	IF InitMqttDone THEN
		pMqttPublishQueue^.AddMessage(
			Payload := REAL_TO_STRING(TOTAL_ACTIVE_ENERGY),
			Topic := CONCAT(CONCAT(MqttPublishTopicPrefix^, MqttPublishTopicSuffix), '/TOTAE' ),
			Qos := MQTT.QoS.ExactlyOnce,
			MqttRetain := FALSE
		);
		pMqttPublishQueue^.AddMessage(
			Payload := REAL_TO_STRING(TOTAL_REACTIVE_ENERGY),
			Topic := CONCAT(CONCAT(MqttPublishTopicPrefix^, MqttPublishTopicSuffix), '/TOTRE' ),
			Qos := MQTT.QoS.ExactlyOnce,
			MqttRetain := FALSE
		);
	END_IF
END_IF
          

METHOD ProcessDataArray
  VAR_INPUT
    Error : POINTER TO BOOL;
    Data : POINTER TO ARRAY[0..124] OF WORD;
  END_VAR
                  IF Error^ THEN
	PubMqttMessage(Suffix := '/availability', Data := 'offline');
ELSE
	PubMqttMessage(Suffix := '/availability', Data := 'online');
END_IF

IF ActiveRtuQuery = 1 THEN
	THIS^.Error1 := Error^;
	THIS^.timerData1.IN := TRUE;
	IF NOT Error^ THEN
		THIS^.VOLTAGE := SwapWordsToReal(Data^[0], Data^[1]);
		THIS^.CURRENT := SwapWordsToReal(Data^[6], Data^[7]);
		THIS^.ACTIVEPOWER := SwapWordsToReal(Data^[12], Data^[13]);
		THIS^.APPARENT_POWER := SwapWordsToReal(Data^[18], Data^[19]);
		THIS^.REACTIVE_POWER := SwapWordsToReal(Data^[24], Data^[25]);
		THIS^.POWER_FACTOR := SwapWordsToReal(Data^[30], Data^[31]);
		THIS^.PHASE_ANGLE := SwapWordsToReal(Data^[36], Data^[37]);
		THIS^.Update1 := TRUE;
	END_IF
ELSIF ActiveRtuQuery = 2 THEN
	THIS^.Error2:= Error^;
	THIS^.timerData2.IN := TRUE;
	IF NOT Error^ THEN		
		THIS^.FREQUENCY := SwapWordsToReal(Data^[0], Data^[1]);
		THIS^.IMPORT_ACTIVE_ENERGY := SwapWordsToReal(Data^[2], Data^[3]);
		THIS^.EXPORT_ACTIVE_ENERGY := SwapWordsToReal(Data^[4], Data^[5]);
		THIS^.IMPORT_REACTIVE_ENERGY := SwapWordsToReal(Data^[6], Data^[7]);
		THIS^.EXPORT_REACTIVE_ENERGY := SwapWordsToReal(Data^[8], Data^[9]);
		THIS^.Update2 := TRUE;
	END_IF
ELSIF ActiveRtuQuery = 3 THEN
	THIS^.Error3 := Error^;
	THIS^.timerData3.IN := TRUE;
	IF NOT Error^ THEN
		THIS^.TOTAL_ACTIVE_ENERGY := SwapWordsToReal(Data^[0], Data^[1]);
		THIS^.TOTAL_REACTIVE_ENERGY := SwapWordsToReal(Data^[2], Data^[3]);
		THIS^.Update3 := TRUE;
	END_IF	
END_IF

ActiveRtuQuery := 0;
ActiveDevice := FALSE;




                
END_METHOD

METHOD InitRS485
  VAR_INPUT
    Data1PollingInterval : TIME;
    Data2PollingInterval : TIME;
    Data3PollingInterval : TIME;
    DeviceAddress : BYTE;
  END_VAR
                  THIS^.timerData1.PT := Data1PollingInterval;
THIS^.timerData2.PT := Data2PollingInterval;
THIS^.timerData3.PT := Data3PollingInterval;

THIS^.Data1RtuQuery.DeviceId := DeviceAddress;
THIS^.Data2RtuQuery.DeviceId := DeviceAddress;
THIS^.Data3RtuQuery.DeviceId := DeviceAddress;

THIS^.timerData1.IN := TRUE;
THIS^.timerData2.IN := TRUE;
THIS^.timerData3.IN := TRUE;

THIS^.InitRS485Done := TRUE;
                
END_METHOD

METHOD InitMqtt
  VAR_INPUT
    MQTTPublishPrefix : POINTER TO STRING;
    pMqttPublishQueue : POINTER TO FB_MqttPublishQueue;
  END_VAR
  VAR
    InstanceNamePt : POINTER TO STRING;
  END_VAR
                  THIS^.pMqttPublishQueue := pMqttPublishQueue;
THIS^.MqttPublishTopicPrefix := MQTTPublishPrefix;

InstanceNamePt := CommonTypesAndFunctions.FindLastDot(ADR(THIS^.InstanceName)) + 1;
THIS^.MqttPublishTopicSuffix := InstanceNamePt^;

THIS^.InitMqttDone := TRUE;
                
END_METHOD

METHOD RequestBusTime : BOOL
                  IF NOT InitRS485Done THEN	
	RequestBusTime := FALSE;	
ELSIF timerData1.Q OR timerData2.Q OR timerData3.Q THEN
	RequestBusTime := TRUE;	
ELSE
	RequestBusTime := FALSE;		
END_IF
                
END_METHOD

METHOD GetRtuQuery : RS485_RtuQuery
                  IF timerData1.Q THEN
	THIS^.timerData1.IN := FALSE;
	THIS^.ActiveRtuQuery := 1;
	GetRtuQuery := THIS^.Data1RtuQuery;
ELSIF timerData2.Q THEN
	THIS^.timerData2.IN := FALSE;
	THIS^.ActiveRtuQuery := 2;
	GetRtuQuery := THIS^.Data2RtuQuery;
ELSIF timerData3.Q THEN
	THIS^.timerData3.IN := FALSE;
	THIS^.ActiveRtuQuery := 3;
	GetRtuQuery := THIS^.Data3RtuQuery;	
END_IF
                
END_METHOD

METHOD PubMqttMessage
  VAR_INPUT
    Suffix : STRING(100);
    Data : STRING(100);
  END_VAR
                  IF InitMqttDone THEN
		pMqttPublishQueue^.AddMessage(
			Payload := Data,
			Topic := CONCAT(CONCAT(MqttPublishTopicPrefix^, MqttPublishTopicSuffix), Suffix ),
			Qos := MQTT.QoS.ExactlyOnce,
			MqttRetain := FALSE
		);
END_IF
                
END_METHOD
END_FUNCTION_BLOCK

{attribute 'reflection'}
FUNCTION_BLOCK FB_RS485_ESERA_1WIRE_GATEWAY_MQTT IMPLEMENTS RS485Device
  VAR
    {attribute 'instance-path'}
    {attribute 'noinit'}
    InstanceName : STRING;  (* object's full instance name *)
    InitRS485Done : BOOL := FALSE;
    DeviceAddress : BYTE;
    OwdDevices : ARRAY[1..30] OF FB_RS485_ESERA_OWD_MQTT;
    ActiveDevice : BOOL := FALSE;
    ActiveOwd : UINT := 0;
    loopCounter : UINT;
    timerData : TON;
  END_VAR

            timerData();

FOR loopCounter := 1 TO 30 DO
	OwdDevices[loopCounter]();
END_FOR
          

METHOD GetRtuQuery : RS485_RtuQuery
                  IF timerData.Q THEN
	THIS^.timerData.IN := FALSE;
	GetRtuQuery := THIS^.OwdDevices[ActiveOwd].GetRtuQuery();	
END_IF
                
END_METHOD

METHOD ProcessDataArray
  VAR_INPUT
    Error : POINTER TO BOOL;
    Data : POINTER TO ARRAY[0..124] OF WORD;
  END_VAR
                  THIS^.OwdDevices[ActiveOwd].ProcessDataArray(
	Data := Data,
	Error := Error
);
THIS^.ActiveOwd := 0;
THIS^.timerData.IN := TRUE;
                
END_METHOD

METHOD RequestBusTime : BOOL
                  IF NOT InitRS485Done OR NOT timerData.Q THEN	
	RequestBusTime := FALSE;
ELSE
	FOR loopCounter := 1 TO 30 DO
		IF OwdDevices[loopCounter].RequestBusTime() AND RequestBusTime = FALSE THEN
			THIS^.ActiveOwd := loopCounter;
			RequestBusTime := TRUE;			
		END_IF
	END_FOR
END_IF
                
END_METHOD

METHOD InitRS485
  VAR_INPUT
    DeviceAddress : BYTE;
  END_VAR
                  THIS^.DeviceAddress := DeviceAddress;
THIS^.timerData.PT := T#250MS;
THIS^.timerData.IN := TRUE;
THIS^.InitRS485Done := TRUE;
                
END_METHOD

METHOD InitMqtt
  VAR_INPUT
    MQTTPublishPrefix : POINTER TO STRING;
    pMqttPublishQueue : POINTER TO FB_MqttPublishQueue;
  END_VAR
  VAR
    InstanceNamePt : POINTER TO STRING;
  END_VAR
                  InstanceNamePt := CommonTypesAndFunctions.FindLastDot(ADR(THIS^.InstanceName)) + 1;

FOR loopCounter := 1 TO 30 DO
		OwdDevices[loopCounter].InitMqtt(
			MQTTPublishPrefix := MQTTPublishPrefix,
			MqttPublishTopicSuffix := InstanceNamePt^,
			pMqttPublishQueue := pMqttPublishQueue
		);
END_FOR
                
END_METHOD

METHOD EnableOwd : BOOL
  VAR_INPUT
    OwdNumber : UINT;
    DataPollingInterval : TIME;
  END_VAR
                  THIS^.OwdDevices[OwdNumber].InitOwd(
	DeviceAddress := THIS^.DeviceAddress,
	OwdNumber := OwdNumber,
	DataPollingInterval := DataPollingInterval
);
                
END_METHOD
END_FUNCTION_BLOCK

FUNCTION_BLOCK FB_RS485_ESERA_OWD_MQTT
  VAR_OUTPUT
    OWD_VOLTAGE : REAL := 0;
    TEMPERATURE : REAL := 0;
    HUMIDITY : REAL := 0;
    DEW_POINT : REAL := 0;
    AIR_QUALITY : REAL := 0;
    BRIGHTNESS : REAL := 0;
    DataAvailable : BOOL := FALSE;
    Error : BOOL := FALSE;
  END_VAR
  VAR
    OwdNumber : UINT;
    InitMqttDone : BOOL;
    MqttPublishTopicPrefix : POINTER TO STRING;
    MqttPublishTopicSuffix : STRING(50);
    pMqttPublishQueue : POINTER TO FB_MqttPublishQueue;
    InitOwdDone : BOOL := FALSE;
    timerData : TON;
    RtuQuery : RS485_RtuQuery := (FunctionCode := 3, ReadAddress := 100, ReadQuantity := 17);
  END_VAR

            timerData();


          

METHOD InitOwd
  VAR_INPUT
    DeviceAddress : BYTE;
    OwdNumber : UINT;
    DataPollingInterval : TIME;
  END_VAR
                  THIS^.RtuQuery.DeviceId := DeviceAddress;
THIS^.RtuQuery.ReadAddress := OwdNumber * 100;
THIS^.timerData.PT := DataPollingInterval;
THIS^.OwdNumber := OwdNumber;

THIS^.timerData.IN := TRUE;

THIS^.InitOwdDone := TRUE;
                
END_METHOD

METHOD InitMqtt
  VAR_INPUT
    MQTTPublishPrefix : POINTER TO STRING;
    MqttPublishTopicSuffix : STRING(255);
    pMqttPublishQueue : POINTER TO FB_MqttPublishQueue;
  END_VAR
                  THIS^.MqttPublishTopicPrefix := MQTTPublishPrefix;
THIS^.MqttPublishTopicSuffix := MqttPublishTopicSuffix;
THIS^.pMqttPublishQueue := pMqttPublishQueue;

THIS^.InitMqttDone := TRUE;
                
END_METHOD

METHOD PubMqttMessage
  VAR_INPUT
    Suffix : STRING(100);
    Data : STRING(100);
  END_VAR
                  IF InitMqttDone THEN
		pMqttPublishQueue^.AddMessage(
			Payload := Data,
			Topic := CONCAT(CONCAT(CONCAT(CONCAT(MqttPublishTopicPrefix^, MqttPublishTopicSuffix), '/OWD/'), UINT_TO_STRING(OwdNumber)), Suffix ),
			Qos := MQTT.QoS.ExactlyOnce,
			MqttRetain := FALSE
		);
END_IF
                
END_METHOD

METHOD ProcessTemperature
  VAR_INPUT
    Data : WORD;
  END_VAR
                  THIS^.TEMPERATURE := WORD_TO_REAL(Data) / 100;
PubMqttMessage(Suffix := '/TEMP', Data := REAL_TO_STRING(TEMPERATURE));
                
END_METHOD

METHOD ProcessOwdVoltage
  VAR_INPUT
    Data : WORD;
  END_VAR
                  THIS^.OWD_VOLTAGE := WORD_TO_REAL(Data) / 100;
PubMqttMessage(Suffix := '/OWDV', Data := REAL_TO_STRING(OWD_VOLTAGE));
                
END_METHOD

METHOD ProcessHumidity
  VAR_INPUT
    Data : WORD;
  END_VAR
                  THIS^.HUMIDITY := WORD_TO_REAL(Data) / 100;
PubMqttMessage(Suffix := '/HUM', Data := REAL_TO_STRING(HUMIDITY));
                
END_METHOD

METHOD ProcessDewPoint
  VAR_INPUT
    Data : WORD;
  END_VAR
                  THIS^.DEW_POINT := WORD_TO_REAL(Data) / 100;
PubMqttMessage(Suffix := '/DEWP', Data := REAL_TO_STRING(DEW_POINT));
                
END_METHOD

METHOD ProcessAirQuality
  VAR_INPUT
    Data : WORD;
  END_VAR
                  THIS^.AIR_QUALITY := WORD_TO_REAL(Data) / 100;
PubMqttMessage(Suffix := '/AIRQ', Data := REAL_TO_STRING(AIR_QUALITY));
                
END_METHOD

METHOD GetRtuQuery : RS485_RtuQuery
                  IF timerData.Q THEN
	THIS^.timerData.IN := FALSE;
	GetRtuQuery := THIS^.RtuQuery;	
END_IF
                
END_METHOD

METHOD ProcessDataArray
  VAR_INPUT
    Error : POINTER TO BOOL;
    Data : POINTER TO ARRAY[0..124] OF WORD;
  END_VAR
                  THIS^.timerData.IN := TRUE;

IF WORD_TO_INT(Data^[12]) <> 0 OR Error^ THEN
	THIS^.Error := TRUE;
	PubMqttMessage(Suffix := '/availability', Data := 'offline');
ELSE 	
	THIS^.Error := FALSE;
	THIS^.DataAvailable := TRUE;
	PubMqttMessage(Suffix := '/availability', Data := 'online');
END_IF

// Data handling
IF NOT Error^ AND WORD_TO_INT(Data^[12]) = 0 THEN
	IF Data^[16] = 11151 OR Data^[16] = 11152 THEN // Temperature, humidity & air quality
		ProcessTemperature(Data^[0]);		
		ProcessOwdVoltage(Data^[2]);
		ProcessHumidity(Data^[4]);
		ProcessDewPoint(Data^[6]);
		ProcessAirQuality(Data^[8]);
	ELSIF Data^[16] = 11102 OR Data^[16] = 11113 OR Data^[16] = 11120 OR Data^[16] = 11148 OR Data^[16] = 11150 OR Data^[16] = 11160 THEN // Temperature, humidity
		ProcessTemperature(Data^[0]);		
		ProcessOwdVoltage(Data^[2]);
		ProcessHumidity(Data^[4]);
		ProcessDewPoint(Data^[6]);
	ELSIF Data^[16] = 11121 OR Data^[16] = 11132 OR Data^[16] = 11134 OR Data^[16] = 11135 THEN // Temperature, humidity, brightness
		ProcessTemperature(Data^[0]);		
		ProcessOwdVoltage(Data^[2]);
		ProcessHumidity(Data^[4]);
		ProcessDewPoint(Data^[6]);
		ProcessBrigthness(Data^[8]);
	ELSIF Data^[16] = 1820  THEN // Temperature DS18B20
        ProcessTemperature(Data^[0]);
	END_IF		
END_IF
                
END_METHOD

METHOD RequestBusTime : BOOL
                  IF NOT InitOwdDone THEN	
	RequestBusTime := FALSE;	
ELSIF timerData.Q THEN
	RequestBusTime := TRUE;
ELSE
	RequestBusTime := FALSE;	
END_IF
                
END_METHOD

METHOD ProcessBrigthness
  VAR_INPUT
    Data : WORD;
  END_VAR
                  THIS^.BRIGHTNESS := WORD_TO_REAL(Data) / 100;
PubMqttMessage(Suffix := '/BNESS', Data := REAL_TO_STRING(BRIGHTNESS));
                
END_METHOD
END_FUNCTION_BLOCK

{attribute 'reflection'}
FUNCTION_BLOCK FB_VIRTUAL_BOOL_MQTT EXTENDS FB_MQTT_BASE IMPLEMENTS MQTT.MQTT_SUBSCRIBE_CALLBACK
  VAR_INPUT
    IN : BOOL;
  END_VAR
  VAR_OUTPUT
    OUT : BOOL;
  END_VAR
  VAR
    {attribute 'instance-path'}
    {attribute 'noinit'}
    InstancePath : STRING;  (* Refelection: object's full instance name *)
    Startup : BOOL := TRUE;
    UpdateFlag : BOOL;
    VirtualMode : VIRTUAL_MODES;
    DefaultValue : BOOL;
    SetDefaultValueStartup : BOOL;
    PublishAtStartup : BOOL;
    UsePersistentAtStartup : BOOL;
    ConfirmReceival : BOOL;
    MqttMessageReceived : BOOL;
    PreviousIn : BOOL;
  END_VAR
  VAR PERSISTENT
    PreviousState : BOOL;  (* To retain output state through powercycles *)
  END_VAR

            IF VirtualMode = VIRTUAL_MODES.Output THEN
	IF (Startup AND PublishAtStartup) OR (UpdateFlag OR IN <> PreviousIn) AND InitMqttDone THEN
	pMqttPublishQueue^.AddMessage(
		Payload := BOOL_TO_STRING(IN),
		Topic := CONCAT(MqttPublishTopicPrefix^, MqttPublishTopicSuffix),
		Qos := MqttQos,
		MqttRetain := MqttRetain
	);
	Startup:=FALSE;
	UpdateFlag := FALSE;
	PreviousIn := IN;
	END_IF
ELSIF VirtualMode = VIRTUAL_MODES.Input THEN
	IF Startup AND SetDefaultValueStartup THEN
		OUT := DefaultValue;
	ELSIF UsePersistentAtStartup THEN
		OUT := PreviousState;
	END_IF	
	
	IF ((Startup AND PublishAtStartup) OR (ConfirmReceival AND MqttMessageReceived)) AND InitMqttDone THEN
	pMqttPublishQueue^.AddMessage(
		Payload := BOOL_TO_STRING(OUT),
		Topic := CONCAT(MqttPublishTopicPrefix^, MqttPublishTopicSuffix),
		Qos := MqttQos,
		MqttRetain := MqttRetain
	);
	Startup:=FALSE;
	MqttMessageReceived := FALSE;
	PreviousState:=OUT;
	END_IF		
	
END_IF
          

METHOD InitMqtt
  VAR_INPUT
    MQTTPublishPrefix : POINTER TO STRING;
    MQTTSubscribePrefix : POINTER TO STRING;
    pMqttPublishQueue : POINTER TO FB_MqttPublishQueue;
    pMqttCallbackCollector : POINTER TO MQTT.CallbackCollector;
    MqttQos : MQTT.QoS;
    MqttRetain : BOOL;
  END_VAR
                  InitMqttDone := TRUE;

SUPER^._InstancePath := THIS^.InstancePath; // Due to reflection its location is important

(*pass trough*)
THIS^.pMqttPublishQueue := pMqttPublishQueue;
THIS^.MqttPublishTopicPrefix:=MQTTPublishPrefix;
THIS^.MQTTSubscribeTopicPrefix:=MQTTSubscribePrefix;
THIS^.pMqttPublishQueue:=pMqttPublishQueue;
THIS^.MqttQos:=MqttQos;
THIS^.MqttRetain:=MqttRetain;


SUPER^.InitBaseMqtt();
pMqttCallbackCollector^.put(instance:= THIS^); // register the FB agains the collector so mqtt events can be received


                
END_METHOD

METHOD PublishReceived : BOOL
  VAR_INPUT
    Data : MQTT.CALLBACK_DATA;  (* Collection of recived Data *)
  END_VAR
                  //first check if Mqtt is initialized and FB in input mode, otherwise do nothing
IF NOT(InitMqttDone) AND VirtualMode <> VIRTUAL_MODES.Input THEN
	//mark the interface call from the collector as done
	PublishReceived := TRUE;
//check if the packet is for this FB
ELSIF CommonTypesAndFunctions.StrEquals(str1:= ADR(MQTTSubscribeTopic), str2:= Data.TopicOut) THEN
	//mark the interface call from the collector as done
	PublishReceived := TRUE;
	//process the data
	IF CommonTypesAndFunctions.StrEquals(str1:= Data.PayloadString, str2:= ADR('TRUE')) THEN
		THIS^.OUT := TRUE;
		MqttMessageReceived := TRUE;
	END_IF
	IF CommonTypesAndFunctions.StrEquals(str1:= Data.PayloadString, str2:= ADR('FALSE')) THEN
		THIS^.OUT := FALSE;
		MqttMessageReceived := TRUE;
	END_IF
END_IF 
                
END_METHOD

METHOD ConfigureFunctionBlockAsVirtualInput : BOOL
  VAR_INPUT
    DefaultValue : BOOL;
    SetDefaultValueStartup : BOOL;
    PublishAtStartup : BOOL;
    UsePersistentAtStartup : BOOL;
    ConfirmReceival : BOOL;
  END_VAR
                  THIS^.DefaultValue:=DefaultValue;
THIS^.SetDefaultValueStartup:=SetDefaultValueStartup;
THIS^.PublishAtStartup:=PublishAtStartup;
THIS^.UsePersistentAtStartup:=UsePersistentAtStartup;
THIS^.ConfirmReceival:=ConfirmReceival;
THIS^.VirtualMode:=VIRTUAL_MODES.Input;
                
END_METHOD

METHOD SetValue : BOOL
  VAR_INPUT
    Value : BOOL;
  END_VAR
                  THIS^.OUT:=Value;
THIS^.UpdateFlag:=TRUE;
                
END_METHOD

METHOD ConfigureFunctionBlockAsVirtualOutput : BOOL
  VAR_INPUT
    PublishAtStartup : BOOL;
  END_VAR
                  THIS^.PublishAtStartup:=PublishAtStartup;
THIS^.VirtualMode:=VIRTUAL_MODES.Output;
                
END_METHOD
END_FUNCTION_BLOCK

{attribute 'reflection'}
FUNCTION_BLOCK FB_VIRTUAL_INT_MQTT EXTENDS FB_MQTT_BASE IMPLEMENTS MQTT.MQTT_SUBSCRIBE_CALLBACK
  VAR_INPUT
    IN : INT;
  END_VAR
  VAR_OUTPUT
    OUT : INT;
  END_VAR
  VAR
    {attribute 'instance-path'}
    {attribute 'noinit'}
    InstancePath : STRING;  (* Refelection: object's full instance name *)
    Startup : BOOL := TRUE;
    UpdateFlag : BOOL;
    VirtualMode : VIRTUAL_MODES;
    DefaultValue : INT;
    SetDefaultValueStartup : BOOL;
    PublishAtStartup : BOOL;
    UsePersistentAtStartup : BOOL;
    ConfirmReceival : BOOL;
    MqttMessageReceived : BOOL;
    PreviousIn : INT;
  END_VAR
  VAR PERSISTENT
    PreviousState : INT;  (* To retain output state through powercycles *)
  END_VAR

            IF VirtualMode = VIRTUAL_MODES.Output THEN
	IF (Startup AND PublishAtStartup) OR (UpdateFlag OR IN <> PreviousIn) AND InitMqttDone THEN
	pMqttPublishQueue^.AddMessage(
		Payload := INT_TO_STRING(IN),
		Topic := CONCAT(MqttPublishTopicPrefix^, MqttPublishTopicSuffix),
		Qos := MqttQos,
		MqttRetain := MqttRetain
	);
	Startup:=FALSE;
	UpdateFlag := FALSE;
	PreviousIn := IN;
	END_IF
ELSIF VirtualMode = VIRTUAL_MODES.Input THEN
	IF Startup AND SetDefaultValueStartup THEN
		OUT := DefaultValue;
	ELSIF UsePersistentAtStartup THEN
		OUT := PreviousState;
	END_IF	
	
	IF ((Startup AND PublishAtStartup) OR (ConfirmReceival AND MqttMessageReceived)) AND InitMqttDone THEN
	pMqttPublishQueue^.AddMessage(
		Payload := INT_TO_STRING(OUT),
		Topic := CONCAT(MqttPublishTopicPrefix^, MqttPublishTopicSuffix),
		Qos := MqttQos,
		MqttRetain := MqttRetain
	);
	Startup:=FALSE;
	MqttMessageReceived := FALSE;
	PreviousState:=OUT;
	END_IF		
	
END_IF
          

METHOD ConfigureFunctionBlockAsVirtualOutput : BOOL
  VAR_INPUT
    PublishAtStartup : BOOL;
  END_VAR
                  THIS^.PublishAtStartup:=PublishAtStartup;
THIS^.VirtualMode:=VIRTUAL_MODES.Output;
                
END_METHOD

METHOD InitMqtt
  VAR_INPUT
    MQTTPublishPrefix : POINTER TO STRING;
    MQTTSubscribePrefix : POINTER TO STRING;
    pMqttPublishQueue : POINTER TO FB_MqttPublishQueue;
    pMqttCallbackCollector : POINTER TO MQTT.CallbackCollector;
    MqttQos : MQTT.QoS;
    MqttRetain : BOOL;
  END_VAR
                  InitMqttDone := TRUE;

SUPER^._InstancePath := THIS^.InstancePath; // Due to reflection its location is important

(*pass trough*)
THIS^.pMqttPublishQueue := pMqttPublishQueue;
THIS^.MqttPublishTopicPrefix:=MQTTPublishPrefix;
THIS^.MQTTSubscribeTopicPrefix:=MQTTSubscribePrefix;
THIS^.pMqttPublishQueue:=pMqttPublishQueue;
THIS^.MqttQos:=MqttQos;
THIS^.MqttRetain:=MqttRetain;


SUPER^.InitBaseMqtt();
pMqttCallbackCollector^.put(instance:= THIS^); // register the FB agains the collector so mqtt events can be received


                
END_METHOD

METHOD PublishReceived : BOOL
  VAR_INPUT
    Data : MQTT.CALLBACK_DATA;  (* Collection of recived Data *)
  END_VAR
                  //first check if Mqtt is initialized and FB in input mode, otherwise do nothing
IF NOT(InitMqttDone) AND VirtualMode <> VIRTUAL_MODES.Input THEN
	//mark the interface call from the collector as done
	PublishReceived := TRUE;
//check if the packet is for this FB
ELSIF CommonTypesAndFunctions.StrEquals(str1:= ADR(MQTTSubscribeTopic), str2:= Data.TopicOut) THEN
	//mark the interface call from the collector as done
	PublishReceived := TRUE;
	//process the data
	IF OSCAT_BASIC.IS_NUM(str:= Data.PayloadString^) THEN
		THIS^.OUT := STRING_TO_INT(Data.PayloadString^);	
		MqttMessageReceived := TRUE;	
	END_IF
END_IF 
                
END_METHOD

METHOD ConfigureFunctionBlockAsVirtualInput : BOOL
  VAR_INPUT
    DefaultValue : INT;
    SetDefaultValueStartup : BOOL;
    PublishAtStartup : BOOL;
    UsePersistentAtStartup : BOOL;
    ConfirmReceival : BOOL;
  END_VAR
                  THIS^.DefaultValue:=DefaultValue;
THIS^.SetDefaultValueStartup:=SetDefaultValueStartup;
THIS^.PublishAtStartup:=PublishAtStartup;
THIS^.UsePersistentAtStartup:=UsePersistentAtStartup;
THIS^.ConfirmReceival:=ConfirmReceival;
THIS^.VirtualMode:=VIRTUAL_MODES.Input;
                
END_METHOD

METHOD SetValue : BOOL
  VAR_INPUT
    Value : INT;
  END_VAR
                  THIS^.OUT:=Value;
THIS^.UpdateFlag:=TRUE;
                
END_METHOD
END_FUNCTION_BLOCK

{attribute 'reflection'}
FUNCTION_BLOCK FB_VIRTUAL_REAL_MQTT EXTENDS FB_MQTT_BASE IMPLEMENTS MQTT.MQTT_SUBSCRIBE_CALLBACK
  VAR_INPUT
    IN : REAL;
  END_VAR
  VAR_OUTPUT
    OUT : REAL;
  END_VAR
  VAR
    {attribute 'instance-path'}
    {attribute 'noinit'}
    InstancePath : STRING;  (* Refelection: object's full instance name *)
    Startup : BOOL := TRUE;
    UpdateFlag : BOOL;
    VirtualMode : VIRTUAL_MODES;
    DefaultValue : REAL;
    SetDefaultValueStartup : BOOL;
    PublishAtStartup : BOOL;
    UsePersistentAtStartup : BOOL;
    ConfirmReceival : BOOL;
    MqttMessageReceived : BOOL;
    PreviousIn : REAL;
  END_VAR
  VAR PERSISTENT
    PreviousState : REAL;  (* To retain output state through powercycles *)
  END_VAR

            IF VirtualMode = VIRTUAL_MODES.Output THEN
	IF (Startup AND PublishAtStartup) OR (UpdateFlag OR IN <> PreviousIn) AND InitMqttDone THEN
	pMqttPublishQueue^.AddMessage(
		Payload := REAL_TO_STRING(IN),
		Topic := CONCAT(MqttPublishTopicPrefix^, MqttPublishTopicSuffix),
		Qos := MqttQos,
		MqttRetain := MqttRetain
	);
	Startup:=FALSE;
	UpdateFlag := FALSE;
	PreviousIn := IN;
	END_IF
ELSIF VirtualMode = VIRTUAL_MODES.Input THEN
	IF Startup AND SetDefaultValueStartup THEN
		OUT := DefaultValue;
	ELSIF UsePersistentAtStartup THEN
		OUT := PreviousState;
	END_IF	
	
	IF ((Startup AND PublishAtStartup) OR (ConfirmReceival AND MqttMessageReceived)) AND InitMqttDone THEN
	pMqttPublishQueue^.AddMessage(
		Payload := REAL_TO_STRING(OUT),
		Topic := CONCAT(MqttPublishTopicPrefix^, MqttPublishTopicSuffix),
		Qos := MqttQos,
		MqttRetain := MqttRetain
	);
	Startup:=FALSE;
	MqttMessageReceived := FALSE;
	PreviousState:=OUT;
	END_IF		
	
END_IF
          

METHOD ConfigureFunctionBlockAsVirtualOutput : BOOL
  VAR_INPUT
    PublishAtStartup : BOOL;
  END_VAR
                  THIS^.PublishAtStartup:=PublishAtStartup;
THIS^.VirtualMode:=VIRTUAL_MODES.Output;
                
END_METHOD

METHOD InitMqtt
  VAR_INPUT
    MQTTPublishPrefix : POINTER TO STRING;
    MQTTSubscribePrefix : POINTER TO STRING;
    pMqttPublishQueue : POINTER TO FB_MqttPublishQueue;
    pMqttCallbackCollector : POINTER TO MQTT.CallbackCollector;
    MqttQos : MQTT.QoS;
    MqttRetain : BOOL;
  END_VAR
                  InitMqttDone := TRUE;

SUPER^._InstancePath := THIS^.InstancePath; // Due to reflection its location is important

(*pass trough*)
THIS^.pMqttPublishQueue := pMqttPublishQueue;
THIS^.MqttPublishTopicPrefix:=MQTTPublishPrefix;
THIS^.MQTTSubscribeTopicPrefix:=MQTTSubscribePrefix;
THIS^.pMqttPublishQueue:=pMqttPublishQueue;
THIS^.MqttQos:=MqttQos;
THIS^.MqttRetain:=MqttRetain;


SUPER^.InitBaseMqtt();
pMqttCallbackCollector^.put(instance:= THIS^); // register the FB agains the collector so mqtt events can be received


                
END_METHOD

METHOD PublishReceived : BOOL
  VAR_INPUT
    Data : MQTT.CALLBACK_DATA;  (* Collection of recived Data *)
  END_VAR
                  //first check if Mqtt is initialized and FB in input mode, otherwise do nothing
IF NOT(InitMqttDone) AND VirtualMode <> VIRTUAL_MODES.Input THEN
	//mark the interface call from the collector as done
	PublishReceived := TRUE;
//check if the packet is for this FB
ELSIF CommonTypesAndFunctions.StrEquals(str1:= ADR(MQTTSubscribeTopic), str2:= Data.TopicOut) THEN
	//mark the interface call from the collector as done
	PublishReceived := TRUE;
	//process the data
	THIS^.OUT := STRING_TO_REAL(Data.PayloadString^);	
	MqttMessageReceived := TRUE;	
END_IF 
                
END_METHOD

METHOD ConfigureFunctionBlockAsVirtualInput : BOOL
  VAR_INPUT
    DefaultValue : REAL;
    SetDefaultValueStartup : BOOL;
    PublishAtStartup : BOOL;
    UsePersistentAtStartup : BOOL;
    ConfirmReceival : BOOL;
  END_VAR
                  THIS^.DefaultValue:=DefaultValue;
THIS^.SetDefaultValueStartup:=SetDefaultValueStartup;
THIS^.PublishAtStartup:=PublishAtStartup;
THIS^.UsePersistentAtStartup:=UsePersistentAtStartup;
THIS^.ConfirmReceival:=ConfirmReceival;
THIS^.VirtualMode:=VIRTUAL_MODES.Input;
                
END_METHOD

METHOD SetValue : BOOL
  VAR_INPUT
    Value : REAL;
  END_VAR
                  THIS^.OUT:=Value;
THIS^.UpdateFlag:=TRUE;
                
END_METHOD
END_FUNCTION_BLOCK

{attribute 'reflection'}
FUNCTION_BLOCK FB_VIRTUAL_STRING_MQTT EXTENDS FB_MQTT_BASE IMPLEMENTS MQTT.MQTT_SUBSCRIBE_CALLBACK
  VAR_INPUT
    IN : STRING;
  END_VAR
  VAR_OUTPUT
    OUT : STRING;
  END_VAR
  VAR
    {attribute 'instance-path'}
    {attribute 'noinit'}
    InstancePath : STRING;  (* Refelection: object's full instance name *)
    Startup : BOOL := TRUE;
    UpdateFlag : BOOL;
    VirtualMode : VIRTUAL_MODES;
    DefaultValue : STRING;
    SetDefaultValueStartup : BOOL;
    PublishAtStartup : BOOL;
    UsePersistentAtStartup : BOOL;
    ConfirmReceival : BOOL;
    MqttMessageReceived : BOOL;
    PreviousIn : STRING;
  END_VAR
  VAR PERSISTENT
    PreviousState : STRING;  (* To retain output state through powercycles *)
  END_VAR

            IF VirtualMode = VIRTUAL_MODES.Output THEN
	IF (Startup AND PublishAtStartup) OR (UpdateFlag OR IN <> PreviousIn) AND InitMqttDone THEN
	pMqttPublishQueue^.AddMessage(
		Payload := IN,
		Topic := CONCAT(MqttPublishTopicPrefix^, MqttPublishTopicSuffix),
		Qos := MqttQos,
		MqttRetain := MqttRetain
	);
	Startup:=FALSE;
	UpdateFlag := FALSE;
	PreviousIn := IN;
	END_IF
ELSIF VirtualMode = VIRTUAL_MODES.Input THEN
	IF Startup AND SetDefaultValueStartup THEN
		OUT := DefaultValue;
	ELSIF UsePersistentAtStartup THEN
		OUT := PreviousState;
	END_IF	
	
	IF ((Startup AND PublishAtStartup) OR (ConfirmReceival AND MqttMessageReceived)) AND InitMqttDone THEN
	pMqttPublishQueue^.AddMessage(
		Payload := OUT,
		Topic := CONCAT(MqttPublishTopicPrefix^, MqttPublishTopicSuffix),
		Qos := MqttQos,
		MqttRetain := MqttRetain
	);
	Startup:=FALSE;
	MqttMessageReceived := FALSE;
	PreviousState:=OUT;
	END_IF		
	
END_IF
          

METHOD InitMqtt
  VAR_INPUT
    MQTTPublishPrefix : POINTER TO STRING;
    MQTTSubscribePrefix : POINTER TO STRING;
    pMqttPublishQueue : POINTER TO FB_MqttPublishQueue;
    pMqttCallbackCollector : POINTER TO MQTT.CallbackCollector;
    MqttQos : MQTT.QoS;
    MqttRetain : BOOL;
  END_VAR
                  InitMqttDone := TRUE;

SUPER^._InstancePath := THIS^.InstancePath; // Due to reflection its location is important

(*pass trough*)
THIS^.pMqttPublishQueue := pMqttPublishQueue;
THIS^.MqttPublishTopicPrefix:=MQTTPublishPrefix;
THIS^.MQTTSubscribeTopicPrefix:=MQTTSubscribePrefix;
THIS^.pMqttPublishQueue:=pMqttPublishQueue;
THIS^.MqttQos:=MqttQos;
THIS^.MqttRetain:=MqttRetain;


SUPER^.InitBaseMqtt();
pMqttCallbackCollector^.put(instance:= THIS^); // register the FB agains the collector so mqtt events can be received


                
END_METHOD

METHOD PublishReceived : BOOL
  VAR_INPUT
    Data : MQTT.CALLBACK_DATA;  (* Collection of recived Data *)
  END_VAR
                  //first check if Mqtt is initialized and FB in input mode, otherwise do nothing
IF NOT(InitMqttDone) AND VirtualMode <> VIRTUAL_MODES.Input THEN
	//mark the interface call from the collector as done
	PublishReceived := TRUE;
//check if the packet is for this FB
ELSIF CommonTypesAndFunctions.StrEquals(str1:= ADR(MQTTSubscribeTopic), str2:= Data.TopicOut) THEN
	//mark the interface call from the collector as done
	PublishReceived := TRUE;
	//process the data
	THIS^.OUT := Data.PayloadString^;	
	MqttMessageReceived := TRUE;
END_IF 
                
END_METHOD

METHOD ConfigureFunctionBlockAsVirtualInput : BOOL
  VAR_INPUT
    DefaultValue : STRING;
    SetDefaultValueStartup : BOOL;
    PublishAtStartup : BOOL;
    UsePersistentAtStartup : BOOL;
    ConfirmReceival : BOOL;
  END_VAR
                  THIS^.DefaultValue:=DefaultValue;
THIS^.SetDefaultValueStartup:=SetDefaultValueStartup;
THIS^.PublishAtStartup:=PublishAtStartup;
THIS^.UsePersistentAtStartup:=UsePersistentAtStartup;
THIS^.ConfirmReceival:=ConfirmReceival;
THIS^.VirtualMode:=VIRTUAL_MODES.Input;
                
END_METHOD

METHOD SetValue : BOOL
  VAR_INPUT
    Value : STRING;
  END_VAR
                  THIS^.OUT:=Value;
THIS^.UpdateFlag:=TRUE;
                
END_METHOD

METHOD ConfigureFunctionBlockAsVirtualOutput : BOOL
  VAR_INPUT
    PublishAtStartup : BOOL;
  END_VAR
                  THIS^.PublishAtStartup:=PublishAtStartup;
THIS^.VirtualMode:=VIRTUAL_MODES.Output;
                
END_METHOD
END_FUNCTION_BLOCK

FUNCTION SwapWordsToReal : REAL
  VAR_INPUT
    wHi : WORD;
    wLo : WORD;
  END_VAR
  VAR
    dwVar : DWORD;
    pt_REAL : POINTER TO REAL;
  END_VAR

            dwVar := SHL(WORD_TO_DWORD(wHi),16) OR WORD_TO_DWORD(wLo);
pt_REAL := ADR(dwVar);
SwapWordsToReal := pt_REAL^;
          
END_FUNCTION

PROGRAM PLC_PRG_MAIN
  VAR
    PLC_Device : FB_PLC_MQTT_DISCOVERY_DEVICE;  (* HOME ASSISTANT DISCOVERY VIA MQTT *)
    FB_DI_PB_001 : FB_INPUT_PUSHBUTTON_MQTT;  (* INPUT FUNCTION BLOCKS *)
    FB_DI_PB_002 : FB_INPUT_PUSHBUTTON_DIMMER_MQTT;
    FB_DO_BIN_001 : FB_OUTPUT_BINARY_MQTT;  (* OUTPUT FUNCTION BLOCKS *)
    FB_DO_BISTABLE_001 : FB_OUTPUT_BISTABLE_MQTT;
    FB_DO_COVER_001 : FB_OUTPUT_COVER_MQTT;  (* COVER FUNCTION BLOCKS *)
    FB_AO_DIMMER_001 : FB_OUTPUT_DIMMER_MQTT;  (* DIMMER FUNCTION BLOCKS *)
    TestOUT : WORD;
    FB_VIRTUAL_INT_001 : FB_VIRTUAL_INT_MQTT;  (* VIRTUAL FUNCTION BLOCKS *)
    FB_VIRTUAL_BOOL_001 : FB_VIRTUAL_BOOL_MQTT;
    FB_VIRTUAL_STRING_001 : FB_VIRTUAL_STRING_MQTT;
    FB_VIRTUAL_REAL_001 : FB_VIRTUAL_REAL_MQTT;
  END_VAR

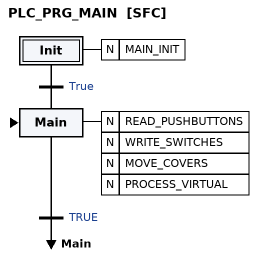
INITIAL_STEP Init:
  MAIN_INIT(N);
END_STEP
TRANSITION FROM Init TO Main
  := True;
END_TRANSITION
STEP Main:
  READ_PUSHBUTTONS(N);
  WRITE_SWITCHES(N);
  MOVE_COVERS(N);
  PROCESS_VIRTUAL(N);
END_STEP
TRANSITION FROM Main TO Main
  := TRUE;
END_TRANSITION

ACTION READ_PUSHBUTTONS:
                      FB_DI_PB_001(PB:= DI_001); (* Provide the input FB the correct phyical input to validate each cyclus *)
FB_DI_PB_002(PB:= DI_002);
                    
END_ACTION

ACTION WRITE_SWITCHES:
                      FB_DO_BIN_001(OUT	=>		DO_001,										(* couple the function block to the physical output *)
	PRIO_HIGH				:=FALSE,  									(* brings the output high regardless of other input values *)
	PRIO_LOW				:=FALSE, 									(* brings the output low regardless of other input values. NOTE: PRIO_HIGH overrules PRIO_LOW input *)
	TOGGLE					:=FB_DI_PB_001.SINGLE 						(* for toggling the output *)	
);

FB_AO_DIMMER_001(
	SINGLE:=FB_DI_PB_001.SINGLE,
	LONG:=FB_DI_PB_001.LONG, 
	P_LONG:=FB_DI_PB_001.P_LONG, 
	Q_OUT => TestOUT,
	SET:=  FB_DI_PB_001.DOUBLE,
	VAL:=125
);

FB_DO_BISTABLE_001();
                    
END_ACTION

ACTION MAIN_INIT:
                      (* MQTT Discovery device*)
PLC_Device.initPlcDevice(
	MqttDiscoveryPrefix := MqttVariables.MqttHADiscoveryPrefix,
	pMqttPublishQueue := ADR(MqttVariables.fbMqttPublishQueue),
	availabilityTopic := MqttVariables.MqttAvailabilityTopic,
	availabilityOnline := MqttVariables.MqttAvailabilityOnlinePayload,
	availabilityOffline := MqttVariables.MqttAvailabilityOfflinePayload
);

(* MQTT logger*)
MqttVariables.MQTT_logger.InitMqtt(
	MQTTPublishPrefix:= ADR(MqttVariables.MqttPubLogPrefix),											
	pMqttPublishQueue := ADR(MqttVariables.fbMqttPublishQueue),				
	MqttQos:=MQTT.QoS.ExactlyOnce, 
	MqttRetain:=FALSE											
);
MqttVariables.MQTT_logger.InitMqttDiscovery(
	Device := ADR(PLC_Device),							(* The device show in Home Assistant *)
);


(* INIT DIGITAL INPUT STUFF *)
FB_DI_PB_001.InitMqtt(
	MQTTPublishPrefix:= ADR(MqttVariables.MqttPushbuttonPrefix),	(* pointer to string prefix for the mqtt publish topic *)
	pMqttPublishQueue := ADR(MqttVariables.fbMqttPublishQueue)		(* pointer to MqttPublishQueue to send a new Mqtt event *)
);

FB_DI_PB_001.InitMqttDiscovery(
	name := 'Button number 001',						(* The name show in Home Assistant frond-end*)
	Device := ADR(PLC_Device),							(* The device show in Home Assistant *)
);

FB_DI_PB_002.InitMqtt(
	MQTTPublishPrefix:= ADR(MqttVariables.MqttPushbuttonPrefix),	
	pMqttPublishQueue := ADR(MqttVariables.fbMqttPublishQueue),
    TRUE,                                                               (* specify whether dimmer value should be outputted on MQTT topic *)
    MQTT.QoS.ExactlyOnce,                                            (* specify the QoS for the dimmer mqtt events (values 0-255) *)    
    5                                                                   (* specify the resolution for the dimmer mqtt events *)    
);


(* ALTER THE DIMMER OUTPUT DEFAULT BEHAVIOR *)
FB_AO_DIMMER_001.ConfigureFunctionBlock(
	T_Debounce:=T#10MS,
	T_Reconfig:=T#10S,
	T_On_Max:=T#0S,
	T_Dimm_Start:=T#400MS,
	T_Dimm:=T#3S,
	Min_On:=50,
	Max_On:=255,
	Soft_Dimm:=TRUE,
	Rst_Out:=FALSE,
	OUT_LinearScaleMin:=11000,
	OUT_LinearScaleMax:=32767
);

(* INIT DMX / ART-NET OUTPUT, OPTIONAL*)
FB_AO_DIMMER_001.InitDmx(
	DmxChannel := 1,							(* The channel *)
	DmxWidth:=1, 								(* Width of DMX channel, 1 or 2, aka 8 or 16 bit *)
	pDmxValues := ADR(DMXVariables.DMX.BUFFER), (* pointer to network buffer *)
	DmxUniverse:=1								(* Universe, but the buffer desides, this is only meta data that ends up in MQTT*)
);

(* INIT HOME ASSISTANT DISCOVERTY*)
FB_AO_DIMMER_001.InitMqttDiscovery(
	name := '001. Office strip cold',					(* The name show in Home Assistant frond-end*)
	Device := ADR(PLC_Device),							(* The device show in Home Assistant *)
);


(* INIT DIGITAL OUTPUT STUFF *)
FB_DO_BISTABLE_001.InitMqtt(
	MQTTPublishPrefix:= ADR(MqttVariables.MqttPubSwitchPrefix),					(* pointer to string prefix for the mqtt publish topic *)
	MQTTSubscribePrefix:= ADR(MqttVariables.MqttSubSwitchPrefix),				(* pointer to string prefix for the mqtt subscribe topic *)
	pMqttPublishQueue := ADR(MqttVariables.fbMqttPublishQueue),					(* pointer to MqttPublishQueue to send a new Mqtt event *)
	pMqttCallbackCollector := ADR(MqttVariables.collector_FB_OUTPUT_SWITCH_MQTT)(* pointer to CallbackCollector to receive Mqtt subscription events *)
);

FB_DO_BISTABLE_001.InitMqttDiscoveryAsLight(
	name := 'light number 1',						(* The name show in Home Assistant frond-end*)
	Device := ADR(PLC_Device),							(* The device show in Home Assistant *)
);

FB_DO_BIN_001.InitMqtt(
	MQTTPublishPrefix:= ADR(MqttVariables.MqttPubSwitchPrefix),					(* pointer to string prefix for the mqtt publish topic *)
	MQTTSubscribePrefix:= ADR(MqttVariables.MqttSubSwitchPrefix),				(* pointer to string prefix for the mqtt subscribe topic *)
	pMqttPublishQueue := ADR(MqttVariables.fbMqttPublishQueue),					(* pointer to MqttPublishQueue to send a new Mqtt event *)
	pMqttCallbackCollector := ADR(MqttVariables.collector_FB_OUTPUT_SWITCH_MQTT)(* pointer to CallbackCollector to receive Mqtt subscription events *)
);

FB_DO_BIN_001.InitMqttDiscoveryAsLight(
	name := 'light number 2',						(* The name show in Home Assistant frond-end*)
	Device := ADR(PLC_Device),							(* The device show in Home Assistant *)
);

(* INIT COVERS STUFF *)
FB_DO_COVER_001.InitMqtt(MQTTPublishPrefix:= ADR(MqttVariables.MqttPubCoverPrefix),	(* pointer to string prefix for the mqtt publish topic *)
	MQTTSubscribePrefix:= ADR(MqttVariables.MqttSubCoverPrefix),					(* pointer to string prefix for the mqtt subscribe topic *)
	pMqttPublishQueue := ADR(MqttVariables.fbMqttPublishQueue),						(* pointer to MqttPublishQueue to send a new Mqtt event *)
	pMqttCallbackCollector := ADR(MqttVariables.collector_FB_OUTPUT_COVER_MQTT)  	(* pointer to CallbackCollector to receive Mqtt subscription events *)
);

FB_DO_COVER_001.initmqttdiscovery(								(*see dimmer for full example *)
	name := 'cover number 001',									(* the name show in home assistant frond-end*)
	device := ADR(PLC_Device),										(* the device show in home assistant *)
);

FB_DO_COVER_001.ConfigureFunctionBlock(
	T_LOCKOUT:=T#1S,											(* delay between change of direction *)
	T_UD:=T#20S													(* run time to move the cover completely up/down *)
);


(* INIT VIRTUAL STUFF *)
FB_VIRTUAL_STRING_001.InitMqtt(MQTTPublishPrefix:= ADR(MqttVariables.MqttPubVirtualPrefix),				
	MQTTSubscribePrefix:= ADR(MqttVariables.MqttSubVirtualPrefix),									
	pMqttPublishQueue := ADR(MqttVariables.fbMqttPublishQueue),						
	pMqttCallbackCollector := ADR(MqttVariables.collector_FB_VIRTUAL_MQTT),
	MqttQos:=MQTT.QoS.ExactlyOnce, 
	MqttRetain:=FALSE									
);
FB_VIRTUAL_STRING_001.ConfigureFunctionBlockAsVirtualInput(DefaultValue:='HelloWorld',SetDefaultValueStartup:=TRUE,PublishAtStartup:=TRUE,UsePersistentAtStartup:=FALSE,ConfirmReceival:=TRUE);


FB_VIRTUAL_INT_001.InitMqtt(MQTTPublishPrefix:= ADR(MqttVariables.MqttPubVirtualPrefix),				
	MQTTSubscribePrefix:= ADR(MqttVariables.MqttSubVirtualPrefix),									
	pMqttPublishQueue := ADR(MqttVariables.fbMqttPublishQueue),						
	pMqttCallbackCollector := ADR(MqttVariables.collector_FB_VIRTUAL_MQTT),
	MqttQos:=MQTT.QoS.ExactlyOnce, 
	MqttRetain:=FALSE												
);
FB_VIRTUAL_INT_001.ConfigureFunctionBlockAsVirtualInput(DefaultValue:=0,SetDefaultValueStartup:=TRUE,PublishAtStartup:=TRUE,UsePersistentAtStartup:=FALSE,ConfirmReceival:=TRUE);
(* FB_VIRTUAL_INT_001.ConfigureFunctionBlockAsVirtualOutput(PublishAtStartup:=TRUE); *)


FB_VIRTUAL_BOOL_001.InitMqtt(MQTTPublishPrefix:= ADR(MqttVariables.MqttPubVirtualPrefix),				
	MQTTSubscribePrefix:= ADR(MqttVariables.MqttSubVirtualPrefix),									
	pMqttPublishQueue := ADR(MqttVariables.fbMqttPublishQueue),						
	pMqttCallbackCollector := ADR(MqttVariables.collector_FB_VIRTUAL_MQTT),
	MqttQos:=MQTT.QoS.ExactlyOnce, 
	MqttRetain:=FALSE											
);
(* FB_VIRTUAL_BOOL_001.ConfigureFunctionBlockAsVirtualInput(DefaultValue:=FALSE,SetDefaultValueStartup:=TRUE,PublishAtStartup:=TRUE,UsePersistentAtStartup:=FALSE); *)
FB_VIRTUAL_BOOL_001.ConfigureFunctionBlockAsVirtualOutput(PublishAtStartup:=TRUE);

FB_VIRTUAL_REAL_001.InitMqtt(MQTTPublishPrefix:= ADR(MqttVariables.MqttPubVirtualPrefix),				
	MQTTSubscribePrefix:= ADR(MqttVariables.MqttSubVirtualPrefix),									
	pMqttPublishQueue := ADR(MqttVariables.fbMqttPublishQueue),						
	pMqttCallbackCollector := ADR(MqttVariables.collector_FB_VIRTUAL_MQTT),
	MqttQos:=MQTT.QoS.ExactlyOnce, 
	MqttRetain:=FALSE												
);
FB_VIRTUAL_REAL_001.ConfigureFunctionBlockAsVirtualInput(DefaultValue:=0.1,SetDefaultValueStartup:=TRUE,PublishAtStartup:=TRUE,UsePersistentAtStartup:=FALSE,ConfirmReceival:=TRUE);
(* FB_VIRTUAL_REAL_001.ConfigureFunctionBlockAsVirtualOutput(PublishAtStartup:=TRUE); *)



MqttVariables.MQTT_logger.send('Init finished', 'MAIN_INIT');


                    
END_ACTION

ACTION MOVE_COVERS:
                      FB_DO_COVER_001(
	TOGGLE:=FB_DI_PB_001.P_LONG,
	MU=>DO_031,
	MD=>DO_032	
);
                    
END_ACTION

ACTION PROCESS_VIRTUAL:
                      
FB_VIRTUAL_BOOL_001();
FB_VIRTUAL_INT_001();
FB_VIRTUAL_STRING_001();
FB_VIRTUAL_REAL_001();
                    
END_ACTION
END_PROGRAM

PROGRAM PLC_PRG_MQTT
  VAR
    MQTTClient : MQTT.MQTTClient;
    MQTT_IN_OUT : MQTT.MQTT_IN_OUT;
    MQTTInfo : MQTT.MQTT_INFO;
    MQTTBirthMessage : MQTT_MESSAGE;
    MQTTBirthHartbeat : OSCAT_BASIC.GEN_PULSE;
    MQTTConnectTrigger : Standard.R_TRIG;
    MQTTPublishBirth : BOOL := TRUE;
    MQTTBirthPublisher : FB_MqttPublishWorker;
    initMqtt : BOOL;  (* variables for MQTT setup *)
    icounter : UDINT;
    ipublishers : UDINT := 40;  (* variables for MQTT publishing *)
    publishers : ARRAY[0..39] OF FB_MqttPublishWorker;
    i : UDINT;  (* variables to work with Mqttbuffer *)
    subscriber_FB_OUTPUT_SWITCH_MQTT : MQTT.MQTTSubscribe;  (* variables for MQTT subscribing *)
    subscriber_FB_OUTPUT_COVER_MQTT : MQTT.MQTTSubscribe;
    subscriber_FB_VIRTUAL_MQTT : MQTT.MQTTSubscribe;
    subscriber_FB_DIMMER_MQTT : MQTT.MQTTSubscribe;
    subscriber_FB_RS485_MQTT : MQTT.MQTTSubscribe;
  END_VAR

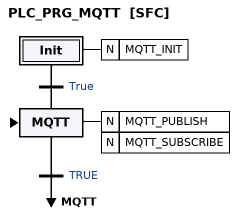
INITIAL_STEP Init:
  MQTT_INIT(N);
END_STEP
TRANSITION FROM Init TO MQTT
  := True;
END_TRANSITION
STEP MQTT:
  MQTT_PUBLISH(N);
  MQTT_SUBSCRIBE(N);
END_STEP
TRANSITION FROM MQTT TO MQTT
  := TRUE;
END_TRANSITION

ACTION MQTT_INIT:
                      
IF NOT initMqtt THEN
	initMqtt := TRUE;
	(* Basic MQTT config *)
	MQTT_IN_OUT.ClientID := MqttVariables.clientID;
	
	(* Set the LWT topic / payload *)
	MQTT_IN_OUT.BuildWillTopicAndMessage := FALSE;
	MQTT_IN_OUT.WillTopicBase := '';
	MQTT_IN_OUT.ClientWillTopic := MqttVariables.MqttAvailabilityTopic;
	MQTT_IN_OUT.ClientWillMessage := MqttVariables.MqttAvailabilityOfflinePayload;
	
	(* Set the birth message *)
	MQTTBirthMessage.Payload := MqttVariables.MqttAvailabilityOnlinePayload;
	MQTTBirthMessage.Topic := MqttVariables.MqttAvailabilityTopic;
	MQTTBirthMessage.Qos := MqttVariables.MQTT_QOS_EXACTLY_ONCE;
	MQTTBirthMessage.MqttRetain := FALSE;
	
	(* Configure the rising edge detector to detect a connect/reconnect to the broker, used for  birth message *)
	MQTTConnectTrigger(CLK := MQTTInfo.MQTT_CONNECTED);
	
	(* Configure the dedicated MQTTBirth publisher *)
	MQTTBirthPublisher.Init(inputMQTT_IN_OUT:= ADR(MQTT_IN_OUT));
	
	(* Configure the pulse generator for the birth message hartbeat *)
	 MQTTBirthHartbeat(ENQ:=TRUE, PTH:=T#0S, PTL:=MqttVariables.MQTTAvailabilityHartbeatTime);
	
	(* INIT MQTT PUBLISH STUFF *)
	FOR icounter := 0 TO (ipublishers-1) DO		
		publishers[icounter].Init(inputMQTT_IN_OUT:= ADR(MQTT_IN_OUT));
	END_FOR 
	
	(* INIT MQTT SUBSCRIBE STUFF *)
	subscriber_FB_OUTPUT_SWITCH_MQTT.SetMqttInOut(MQTT_IN_OUT:= MQTT_IN_OUT);	
	subscriber_FB_OUTPUT_COVER_MQTT.SetMqttInOut(MQTT_IN_OUT:= MQTT_IN_OUT);
	subscriber_FB_VIRTUAL_MQTT.SetMqttInOut(MQTT_IN_OUT:= MQTT_IN_OUT);	
	subscriber_FB_DIMMER_MQTT.SetMqttInOut(MQTT_IN_OUT:= MQTT_IN_OUT);
	subscriber_FB_RS485_MQTT.SetMqttInOut(MQTT_IN_OUT:= MQTT_IN_OUT);
END_IF


                    
END_ACTION

ACTION MQTT_PUBLISH:
                      (* set user led green if connected to MQTT broker, flashing red if not *)
(* é!COCKPIT version *)
(* LED_1_BrokerStatus(eID:=eLedID.AppLED_1, xOpen:=TRUE );
IF(MQTTClient.connected) THEN
	LED_1_BrokerStatus.SetStatic(eLedColor.Green);
ELSE
	LED_1_BrokerStatus.SetFlash(T#1S,eLedColor.Red, eLedColor.Off);  
END_IF *)
(* Codesys 3S version *)
(*
IF MQTTClient.connected THEN
     PFC.SetLed(which:=PFC.LED.U1, how:=PFC.LedState.STATIC_GRN);
ELSE
     PFC.SetLed(which:=PFC.LED.U1, how:=PFC.LedState.BLINK_RED);
END_IF 
*)

(* allow the rising edge detector to detect a connect/reconnect to the broker, used for  birth message *)
MQTTConnectTrigger(CLK := MQTTInfo.MQTT_CONNECTED);

(* allow the pulse generator to generate a pulse, used for birth message hartbeat *)
MQTTBirthHartbeat(ENQ:=TRUE, PTH:=T#0S, PTL:=MqttVariables.MQTTAvailabilityHartbeatTime);

(* Check if this is a new connection due to startup or connection issues *)
IF initMqtt AND (MQTTConnectTrigger.Q OR MQTTBirthHartbeat.Q) THEN
	MQTTPublishBirth := TRUE;
END_IF

(* On connect or reconnect publish a birth message using the dedicated birth publisher *)
IF MQTTPublishBirth THEN
	MQTTBirthPublisher.PublishMessage(MqttMessage := MQTTBirthMessage);
	MQTTPublishBirth:=FALSE;
END_IF


(* Check if Mqtt is initialized AND if there are elements on the queue to process AND if a MQTTbirthmessage has been published successfully *)
IF initMqtt AND NOT(MqttVariables.fbMqttPublishQueue.EMPTY) AND MQTTPublishBirth = FALSE AND MQTTBirthPublisher.SendDone THEN	
	(* Loop through all free publishers untill there are no more elements in the queue or no more free publishers *)
	FOR i:=0 TO (ipublishers-1) DO			
		(* use the publishers that are free  *)
		IF publishers[i].SendDone AND NOT(MqttVariables.fbMqttPublishQueue.EMPTY) THEN	
			(* Pass message from the queue to a publisher *)
			publishers[i].PublishMessage(MqttMessage:= MqttVariables.fbMqttPublishQueue.GetMessage());
		ELSIF MqttVariables.fbMqttPublishQueue.EMPTY THEN
			(* Queue is empty, jump out of the for loop	*)
			EXIT;	
		END_IF
	END_FOR
END_IF


(* If MQTT is initialized, let the MqttPublishWorkers do their work *)
IF initMqtt THEN	
	MQTT_IN_OUT.clientFB(
		MQTT_IN_OUT:= MQTT_IN_OUT, 
		ENABLE:= TRUE, 
		URL:= MQttVariables.broker, 
		TIMEOUT:= T#1S, 
		TLS:= FALSE);		
		
	MQTTBirthPublisher();
	
	FOR i := 0 TO (ipublishers-1) DO
  		publishers[i]();
	END_FOR

END_IF

                    
END_ACTION

ACTION MQTT_SUBSCRIBE:
                      (* If MQTT is initialized, let the subscriber(s) do its work *)
IF initMqtt THEN
	
	MQTT_IN_OUT.clientFB(
		MQTT_IN_OUT:= MQTT_IN_OUT, 
		ENABLE:= TRUE, 
		URL:= MqttVariables.broker, 
		TIMEOUT:= T#1S, 
		TLS:= FALSE);

	subscriber_FB_OUTPUT_SWITCH_MQTT(
		Subscribe:= TRUE, 
		Topic:= ADR(MqttVariables.MqttSubSwitchTopic), 
		QoSSubscribe:= MqttVariables.MQTT_QOS_EXACTLY_ONCE, 
		ExpectingString:= TRUE, 
		Callback:= MqttVariables.collector_FB_OUTPUT_SWITCH_MQTT,
	);	
	subscriber_FB_OUTPUT_COVER_MQTT(
		Subscribe:= TRUE, 
		Topic:= ADR(MqttVariables.MqttSubCoverTopic), 
		QoSSubscribe:= MqttVariables.MQTT_QOS_EXACTLY_ONCE, 
		ExpectingString:= TRUE, 
		Callback:= MqttVariables.collector_FB_OUTPUT_COVER_MQTT,
	);	
	subscriber_FB_VIRTUAL_MQTT(
		Subscribe:= TRUE, 
		Topic:= ADR(MqttVariables.MqttSubVirtualTopic), 
		QoSSubscribe:= MqttVariables.MQTT_QOS_EXACTLY_ONCE, 
		ExpectingString:= TRUE, 
		Callback:= MqttVariables.collector_FB_VIRTUAL_MQTT,
	);
	subscriber_FB_DIMMER_MQTT(
		Subscribe:= TRUE, 
		Topic:= ADR(MqttVariables.MqttSubDimmerTopic), 
		QoSSubscribe:= MqttVariables.MQTT_QOS_EXACTLY_ONCE, 
		ExpectingString:= TRUE, 
		Callback:= MqttVariables.collector_FB_DIMMER_MQTT,
	);
	subscriber_FB_RS485_MQTT(
		Subscribe:= TRUE, 
		Topic:= ADR(MqttVariables.MqttSubRS485Topic), 
		QoSSubscribe:= MqttVariables.MQTT_QOS_EXACTLY_ONCE,
		ExpectingString:= TRUE, 
		Callback:= MqttVariables.collector_FB_RS485_MQTT,
	);
END_IF
                    
END_ACTION
END_PROGRAM

PROGRAM PLC_PRG_RS485
  VAR
    ModbusMaster : WagoAppPlcModbus.FbMbMasterSerial := (xConnect := TRUE, udiBaudrate := 9600, usiDataBits := 8, eParity := WagoTypesCom.eTTYParity.None, eStopBits := WagoTypesCom.eTTYStopBits.One, eHandshake := WagoTypesCom.eTTYHandshake.None, ePhysical := WagoTypesCom.eTTYPhysicalLayer.RS485_HalfDuplex, eFrameType := eMbFrameType.RTU, tTimeOut := TIME#500ms);  (* CODESYS 3S Version version xComPortOpen : BOOL; xComPortError : BOOL; rtsResult : RTS_IEC_RESULT; stComPortSettings : SysCom.SysComSettings :=( ulBaudrate :=9600, byParity := 0, byStopBits:=1, ulTimeout :=500, ulBufferSize :=256, sPort:=SYS_COM_PORTS.SYS_COMPORT1 ); hComPort : RTS_IEC_HANDLE; awReadBuffer : ARRAY[0..124] OF WORD; awWriteBuffer : ARRAY[0..124] OF WORD; fbModbusRequest : IoDrvModbus.ModbusRequest2; eComError : IoDrvModbus.MB_ErrorCodes; é!COCKPIT version *)
    RtuQuery : WagoAppPlcModbus.typMbQuery;
    RtuResponse : WagoAppPlcModbus.typMbResponse;
    Trigger : BOOL := FALSE;  (* Shared variables for é!COCKPIT and CODESYS 3S Version *)
    InitRS485 : BOOL := FALSE;
    ActiveRtuQuery : RS485_RtuQuery;
    RS485BusController : FB_RS485_BUSCONTROLLER;
    FB_RS485_EASTRON_SDM220_1 : FB_RS485_EASTRON_SDM220_MQTT;  (* RS485 *)
    FB_RS485_ESERA_1WIRE_GATEWAY_MQTT_HOME : FB_RS485_ESERA_1WIRE_GATEWAY_MQTT;
    FB_RS485_DUCO_DUCOBOX_HOME : FB_RS485_DUCO_DUCOBOX_MQTT;
  END_VAR

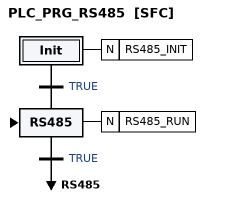
INITIAL_STEP Init:
  RS485_INIT(N);
END_STEP
TRANSITION FROM Init TO RS485
  := TRUE;
END_TRANSITION
STEP RS485:
  RS485_RUN(N);
END_STEP
TRANSITION FROM RS485 TO RS485
  := TRUE;
END_TRANSITION

ACTION RS485_RUN:
                      (* CODESYS 3S Version version*)
(*
IF(NOT xComPortOpen AND NOT xComPortError) THEN
    hComPort := SysCom.SysComOpen2( pSettings := ADR(stComPortSettings), pSettingsEx := 0, pResult := ADR(rtsResult));     
    xComPortError := (hComPort = RTS_INVALID_HANDLE OR rtsResult <> 0);
    xComPortOpen := NOT xComPortError;
END_IF


IF xComPortOpen THEN
	fbModbusRequest.modbusCommand.uiFunctionCode := RS485BusController.ActiveRtuQuery.FunctionCode;
    fbModbusRequest.modbusCommand.uiReadOffset := RS485BusController.ActiveRtuQuery.ReadAddress;	
    fbModbusRequest.modbusCommand.uiReadLen :=RS485BusController.ActiveRtuQuery.ReadQuantity;	   
    fbModbusRequest.pRecvData := ADR(awReadBuffer);
    fbModbusRequest.pSendData := ADR(awWriteBuffer);        
    fbModbusRequest.tResponseTimeout := T#1S;
	fbModbusRequest.transmission := MB_Transmission.RTU;
    fbModbusRequest(
        hComPort := hComPort,
        xExecute := Trigger,
        usiSlaveAddr := RS485BusController.ActiveRtuQuery.DeviceId,		
        byModbusError => eComError);
		
END_IF
*)
	
(* é!COCKPIT version*)
RtuQuery.bUnitId := RS485BusController.ActiveRtuQuery.DeviceId;	
RtuQuery.bFunctionCode := RS485BusController.ActiveRtuQuery.FunctionCode;	
RtuQuery.uiReadAddress := RS485BusController.ActiveRtuQuery.ReadAddress;	
RtuQuery.uiReadQuantity := RS485BusController.ActiveRtuQuery.ReadQuantity;
ModbusMaster(
	I_Port := IoConfig_Globals.COM1,
	utQuery:= RtuQuery,
	xTrigger := Trigger,
	utResponse:= RtuResponse);


(* Shared variables for é!COCKPIT and CODESYS 3S Version *)
RS485BusController();

(* RS485 devices *)
FB_RS485_EASTRON_SDM220_1();
FB_RS485_ESERA_1WIRE_GATEWAY_MQTT_HOME();
FB_RS485_DUCO_DUCOBOX_HOME();
                    
END_ACTION

ACTION RS485_INIT:
                      IF NOT InitRS485 THEN
	InitRS485 := TRUE;

(* INIT RS485 BUS CONTROLLER; CODESYS 3S Version version *)
(*
RS485BusController.Init(
	StartupDelay := T#5S,				(* Time to wait after startup to start using the bus, prevents boot delay issues when RS485 are not ready yet on startup *)		
	SilenceTime := T#50MS,				(* Silence time between two requests, important to not get faulty data on bus *)
	BusTrigger := ADR(Trigger),			(* Pointer to the bool used to initiate bus requests *)
	BusData := ADR(awReadBuffer),		(* Pointer to the array containing the bus response data *)
	BusError := ADR(xComPortError)		(* Pointer to the bus error bool *)
);
*)

(* INIT RS485 BUS CONTROLLER; é!COCKPIT version *)
RS485BusController.Init(
	StartupDelay := T#5S,				(* Time to wait after startup to start using the bus, prevents boot delay issues when RS485 are not ready yet on startup *)		
	SilenceTime := T#50MS,				(* Silence time between two requests, important to not get faulty data on bus *)
	BusTrigger := ADR(Trigger),			(* Pointer to the bool used to initiate bus requests *)
	BusData := ADR(RtuResponse.awData),	(* Pointer to the array containing the bus response data *)
	BusError := ADR(ModbusMaster.xError)(* Pointer to the bus error bool *)
);

RS485BusController.RegisterDevice(device := FB_RS485_EASTRON_SDM220_1);
RS485BusController.RegisterDevice(device := FB_RS485_ESERA_1WIRE_GATEWAY_MQTT_HOME);
RS485BusController.RegisterDevice(device := FB_RS485_DUCO_DUCOBOX_HOME);

(* INIT RS485 DEVICE STUFF *)
FB_RS485_EASTRON_SDM220_1.InitRS485(
	Data1PollingInterval := T#10S,		(* Polling interval for data array 1 *)				
	Data2PollingInterval := T#20S,		(* Polling interval for data array 2 *)			
	Data3PollingInterval := T#30S,		(* Polling interval for data array 3 *)			
	DeviceAddress := 1					(* Device address of the modbus device *)			
);

FB_RS485_EASTRON_SDM220_1.InitMqtt(
	MQTTPublishPrefix:= ADR(MqttVariables.MqttPubRS485Prefix),						(* pointer to string prefix for the mqtt publish topic *)
	pMqttPublishQueue := ADR(MqttVariables.fbMqttPublishQueue)		(* pointer to MqttPublishQueue to send a new Mqtt event *)
);

FB_RS485_ESERA_1WIRE_GATEWAY_MQTT_HOME.InitRS485(
	DeviceAddress := 2
);

FB_RS485_ESERA_1WIRE_GATEWAY_MQTT_HOME.InitMqtt(
	MQTTPublishPrefix:= ADR(MqttVariables.MqttPubRS485Prefix),	
	pMqttPublishQueue := ADR(MqttVariables.fbMqttPublishQueue)
);

(* ENABLE OWD DEVICES ON ESARE GATEWAY *)
FB_RS485_ESERA_1WIRE_GATEWAY_MQTT_HOME.EnableOwd(
	OwdNumber := 1,
	DataPollingInterval := T#2M
);

FB_RS485_ESERA_1WIRE_GATEWAY_MQTT_HOME.EnableOwd(
	OwdNumber := 2,
	DataPollingInterval := T#2M
);

FB_RS485_DUCO_DUCOBOX_HOME.InitRS485(
	DataPollingInterval := T#3S,		(* Polling interval for data array *)				
	DeviceAddress := 3,					(* Device address of the modbus device *)
);

// Nodes: valves for example
FB_RS485_DUCO_DUCOBOX_HOME.AddNode(
	DataPollingInterval := T#15S
);
FB_RS485_DUCO_DUCOBOX_HOME.AddNode(
	DataPollingInterval := T#15S
);

FB_RS485_DUCO_DUCOBOX_HOME.InitMqtt(
	MQTTPublishPrefix:= ADR(MqttVariables.MqttPubRS485Prefix),
	MQTTSubscribePrefix:= ADR(MqttVariables.MqttSubRS485Prefix),
	pMqttPublishQueue := ADR(MqttVariables.fbMqttPublishQueue),	
	pMqttCallbackCollector := ADR(MqttVariables.collector_FB_RS485_MQTT)
);


END_IF
                    
END_ACTION
END_PROGRAM

PROGRAM DMX_SEND
  VAR
    Universe : INT := 1;
    IP_CONTROL2 : oscat_network.IP_CONTROL2;
    IP_C : oscat_network.IP_C;
    S_BUF1 : oscat_network.NETWORK_BUFFER_SHORT;
    R_BUF1 : oscat_network.NETWORK_BUFFER_SHORT;
    error_send : BOOL := FALSE;
    i : INT;
    init : BOOL;
    start : INT;
    size : INT;
    LED_1_BrokerStatus : FbAppLED;
    Step : INT := 0;
  END_VAR

                  IF init = FALSE THEN
	init := TRUE;
	//https://art-net.org.uk/how-it-works/streaming-packets/artdmx-packet-definition/
	(* Write DMX header character in the buffer *) 
	S_BUF1.BUFFER [0]:= BYTE#16#41; // A
	S_BUF1.BUFFER [1]:= BYTE#16#72; // R	
	S_BUF1.BUFFER [2]:= BYTE#16#74; // T
	S_BUF1.BUFFER [3]:= BYTE#16#2D; // -
	S_BUF1.BUFFER [4]:= BYTE#16#4E; // N
	S_BUF1.BUFFER [5]:= BYTE#16#65; // E
	S_BUF1.BUFFER [6]:= BYTE#16#74; // T
	S_BUF1.BUFFER [7]:= BYTE#16#00; // 0 zero
	
	S_BUF1.BUFFER [8]:= BYTE#16#00;	// Opcode ArtDMX (0x5000) little endian
	S_BUF1.BUFFER [9]:= BYTE#16#50; // Opcode ArtDMX (0x5000) little endian
	
	S_BUF1.BUFFER [10]:= BYTE#16#00; // Protocol Version Hi (0)
	S_BUF1.BUFFER [11]:= BYTE#16#0E; // Protocol Version Lo (14)
	
	S_BUF1.BUFFER [12]:= BYTE#16#00; // Sequence
	S_BUF1.BUFFER [13]:= BYTE#16#00; // Physical
	
	S_BUF1.BUFFER [16]:= BYTE#16#02; // Length Hi
	S_BUF1.BUFFER [17]:= BYTE#16#00; // Length Lo (2 to 512, even)
	(* the DMX channels that are next have already been written to the buffer *) 
	
	IF Universe = 1 THEN
		S_BUF1.BUFFER [14]:= BYTE#16#01; // Universe little endian
		S_BUF1.BUFFER [15]:= BYTE#16#00; // Universe little endian
	END_IF
	IF Universe = 2 THEN
		S_BUF1.BUFFER [14]:= BYTE#16#02; // Universe little endian
		S_BUF1.BUFFER [15]:= BYTE#16#00; // Universe little endian
	END_IF
END_IF;


size := 512+18;
FOR i:= 0 TO size DO (* check whether the DMX values ​​in the global variable have changed *)
	// i+2 is strange, buffers are not the same, its often offset with 2 sometimes by 1, todo
	IF S_BUF1.BUFFER[i+18] <> DMXVariables.DMX.BUFFER[i+2] THEN
   		S_BUF1.BUFFER[i+18]:= DMXVariables.DMX.BUFFER[i+2];
		Step := 1;
	END_IF
END_FOR

S_BUF1.BUFFER [17]:= S_BUF1.BUFFER [17]; // low...
DMXVariables.DMX.BUFFER[0] := DMXVariables.DMX.BUFFER[0];
S_BUF1.BUFFER [18]:= S_BUF1.BUFFER [18];
DMXVariables.DMX.BUFFER[1] := DMXVariables.DMX.BUFFER[1];
S_BUF1.BUFFER [19]:= S_BUF1.BUFFER [19];
DMXVariables.DMX.BUFFER[2] := DMXVariables.DMX.BUFFER[2];
S_BUF1.BUFFER [20]:= S_BUF1.BUFFER [20];
DMXVariables.DMX.BUFFER[3] := DMXVariables.DMX.BUFFER[3];


CASE Step OF
	0:
		//passive
	
	1:
		IP_C.C_MODE := 1; (* Mode: UDP+ACTIVE+Port+IP *)
		IP_C.C_ENABLE := TRUE; (* Release connection *)
		IP_C.TIME_RESET := TRUE; (*Reset TIME monitoring * *)
		IP_C.R_OBSERVE := TRUE; (* Monitor data receive *)
		R_BUF1.SIZE:= 0; (* Reset Home length *)
		IP_C.C_IP:= oscat_network.IP4_DECODE (DMXVariables.IP);
		IP_C.C_PORT:= WORD#6454;
		
		S_BUF1.SIZE := size;
		Step:=2;
		
	2:
		IP_CONTROL2 (TIME_OUT:= T#1S, IP_C:= IP_C, S_BUF:= S_BUF1, R_BUF:= R_BUF1);
		
		IF IP_C.ERROR <> 0  THEN
			Step:=666;
		END_IF
	666:
		LED_1_BrokerStatus(eID:=eLedID.AppLED_1, xOpen:=TRUE );
		LED_1_BrokerStatus.SetFlash(T#2S,eLedColor.Red, eLedColor.Off);
		IF IP_C.ERROR = 33554432  THEN
		MqttVariables.MQTT_logger.send(CONCAT('ERROR|DMX has a connection error ', DWORD_TO_STRING(IP_C.ERROR)));
		
		END_IF;
		
		error_send := TRUE;
		R_BUF1.SIZE := 0;
		IP_C.C_ENABLE:= FALSE; (* Enable connection establishment *) 
		IP_C.TIME_RESET:= FALSE;
		init:=FALSE;
	ELSE
	  Step := 0;
END_CASE



// Check IP_C1.error
// 33554432 = 0x02000000
// Initialization of the socket interface failed (only WinNT).
// code = 0x 02 00 00 00 (hexadecimal)
//           !   !    ! 
//           !   !    Receive error 
//           !   Send error
//           Connect error

                
END_PROGRAM

PROGRAM PRG_PING_DMX
  VAR
    PingTime : UDINT;
    DMXnodeReachable : UDINT;
    LED_1_BrokerStatus : FbAppLED;
  END_VAR

                  (* Ping the DMX artNet node *)
DMXnodeReachable := SysSockPing(szIPAddress:=DMXVariables.IP, ulTimeout:=500, pulReplyTime:= ADR(PingTime));

IF DMXnodeReachable = 0 THEN
	LED_1_BrokerStatus.SetStatic(eLedColor.Green);
// 	MqttVariables.MQTT_logger.send('DMX ping OK');
ELSIF DMXnodeReachable = 5 THEN
	LED_1_BrokerStatus.SetFlash(T#1S,eLedColor.Red, eLedColor.Off);
	MqttVariables.MQTT_logger.send('DMX ping Error');
END_IF
                
END_PROGRAM

CONFIGURATION Application
  RESOURCE HomeAutomation ON PLC
    {attribute 'qualified_only'}
    VAR_GLOBAL  (* MqttVariables *)
      clientID : STRING := 'PLC-House';  (* Broker setup *)
      broker : STRING := '192.168.1.52:1883';
      fbMqttPublishQueue : FB_MqttPublishQueue;  (* use the below for username password authentication to broker broker :STRING:='user:password@192.168.1.36:1883'; Shared Variables for MQTT publish communication *)
      collector_FB_OUTPUT_SWITCH_MQTT : MQTT.CallbackCollector;  (* Shared Variables for MQTT subscribe communication *)
      collector_FB_OUTPUT_COVER_MQTT : MQTT.CallbackCollector;
      collector_FB_VIRTUAL_MQTT : MQTT.CallbackCollector;
      collector_FB_DIMMER_MQTT : MQTT.CallbackCollector;
      collector_FB_MQTT_LOG : MQTT.CallbackCollector;
      collector_FB_RS485_MQTT : MQTT.CallbackCollector;
      MQTT_logger : FB_MQTT_LOG;
      MQTT_QOS_EXACTLY_ONCE : MQTT.QoS := MQTT.QoS.ExactlyOnce;  (* QOS Constants *)
      MqttMain : STRING(16) := 'Devices/';  (* Topics *)
      MqttType : STRING(16) := 'PLC/';
      MqttDevice : STRING(16) := 'House/';
      MqttBaseTopic : STRING(100) := 'CONCAT(CONCAT(MqttMain, MqttType), MqttDevice)';  (* e.g. Devices/PLC/House *)
      MqttAvailabilityTopic : STRING(100) := 'CONCAT(MqttBaseTopic, 'availability')';
      MqttAvailabilityOnlinePayload : STRING(20) := 'online';
      MqttAvailabilityOfflinePayload : STRING(20) := 'offline';
      MQTTAvailabilityHartbeatTime : TIME := TIME#5s0ms;
      MqttPubLogPrefix : STRING(100) := 'CONCAT(MqttBaseTopic, 'logger/')';
      MqttHADiscoveryPrefix : STRING(16) := 'homeassistant/';
      MqttPushbuttonPrefix : STRING(100) := 'CONCAT(MqttBaseTopic, 'Out/DigitalInputs/Pushbuttons/')';  (* FB Topics *)
      MqttPubSwitchPrefix : STRING(100) := 'CONCAT(MqttBaseTopic, 'Out/DigitalOutputs/')';
      MqttSubSwitchPrefix : STRING(100) := 'CONCAT(MqttBaseTopic, 'In/DigitalOutputs/')';
      MqttPubCoverPrefix : STRING(100) := 'CONCAT(MqttBaseTopic, 'Out/Covers/')';
      MqttSubCoverPrefix : STRING(100) := 'CONCAT(MqttBaseTopic, 'In/Covers/')';
      MqttPubDimmerPrefix : STRING(100) := 'CONCAT(MqttBaseTopic, 'Out/Dimmers/')';
      MqttSubDimmerPrefix : STRING(100) := 'CONCAT(MqttBaseTopic, 'In/Dimmers/')';
      MqttPubVirtualPrefix : STRING(100) := 'CONCAT(MqttBaseTopic, 'Out/Virtuals/')';
      MqttSubVirtualPrefix : STRING(100) := 'CONCAT(MqttBaseTopic, 'In/Virtuals/')';
      MqttPubRS485Prefix : STRING(100) := 'CONCAT(MqttBaseTopic, 'Out/RS485/')';
      MqttSubRS485Prefix : STRING(100) := 'CONCAT(MqttBaseTopic, 'In/RS485/')';
      MqttSubSwitchTopic : STRING(100) := 'CONCAT(MqttSubSwitchPrefix, '+')';  (* Wildcard subscriptions *)
      MqttSubCoverTopic : STRING(100) := 'CONCAT(MqttSubCoverPrefix, '+')';
      MqttSubVirtualTopic : STRING(100) := 'CONCAT(MqttSubVirtualPrefix, '+')';
      MqttSubDimmerTopic : STRING(100) := 'CONCAT(MqttSubDimmerPrefix, '#')';
      MqttSubRS485Topic : STRING(100) := 'CONCAT(MqttSubRS485Prefix, '#')';
    END_VAR
    {attribute 'qualified_only'}
    VAR_GLOBAL  (* DMXVariables *)
      IP : STRING := '10.1.1.4';  (* unicast: 10.1.1.4 multicast: 10.1.1.255 broadcast: 255.255.255.255 *)
      DMX : oscat_network.NETWORK_BUFFER_SHORT;
    END_VAR
    TASK MainTask(INTERVAL := T#50ms, PRIORITY := 4);
    TASK MqttCommunication(PRIORITY := 5);
    TASK RS485(INTERVAL := T#200ms, PRIORITY := 15);
    TASK Ping(INTERVAL := T#10000ms, PRIORITY := 4);
    PROGRAM PLC_PRG_MAIN WITH MainTask : PLC_PRG_MAIN;
    PROGRAM PLC_PRG_MQTT WITH MqttCommunication : PLC_PRG_MQTT;
    PROGRAM DMX_SEND WITH MqttCommunication : DMX_SEND;
    PROGRAM PLC_PRG_RS485 WITH RS485 : PLC_PRG_RS485;
    PROGRAM PRG_PING_DMX WITH Ping : PRG_PING_DMX;
  END_RESOURCE
END_CONFIGURATION
